Fanuc KAREL source: kc00046.KL

-- PROVISIONAL review KL for V1013-1; original PC SHA256 e5ba4c0fdcc468c6c3b141b72aed118f3ec6d75b333a8cbe41f2f463c03bafcd
-- Incomplete behavior may be omitted. Consult companion uncertainty JSON. Do not deploy.
PROGRAM KC00046
%NOLOCKGROUP
BEGIN
  -- UNRESOLVED_PC offsets 5-27; opcodes 27,22,22,22,31
  -- UNRESOLVED_PC offsets 32-36; opcodes 7F
END KC00046
